(*
SPDX-FileCopyrightText: c 2026 Oleksandr Tiutyk <trofimich@gmail.com>
SPDX-License-Identifier: MIT
License: https://opensource.org/license/mit
*)

(*!
<summary>Checks trimming direction, custom characters and complete removal.</summary>
<description>
Uses one task and stays at a stable address while assertions are bound to this instance.
</description>
*)

{attribute 'no_assign'}
{attribute 'no_explicit_call' := 'do not call this function block directly'}
FUNCTION_BLOCK StringTrimTest EXTENDS TOF_Testing.SingleCycleTest
VAR_STAT
	{attribute 'hide'}
	_ClassName : STRING := __POUNAME();
END_VAR

(*!
<summary>Checks trimming direction, custom characters and complete removal.</summary>
*)
METHOD PROTECTED ExecuteTest
VAR
	text : STRING;
END_VAR
text := '  123   ';
TOF_Core.Strings.TrimChar(stringToTrim := text, trimMode := TOF_Core.TRIM_MODE.LEFT_AND_RIGHT);
Assert.ThatBool(
	actual := text = '123',
	message := "TrimChar must apply LEFT_AND_RIGHT exactly"
).IsTrue();

text := '  123   ';
TOF_Core.Strings.TrimChar(stringToTrim := text, trimMode := TOF_Core.TRIM_MODE.LEFT);
Assert.ThatBool(
	actual := text = '123   ',
	message := "TrimChar must apply LEFT exactly"
).IsTrue();

text := '  123   ';
TOF_Core.Strings.TrimChar(stringToTrim := text, trimMode := TOF_Core.TRIM_MODE.RIGHT);
Assert.ThatBool(
	actual := text = '  123',
	message := "TrimChar must apply RIGHT exactly"
).IsTrue();

text := '**a*b**';
TOF_Core.Strings.TrimChar(stringToTrim := text, trimMode := TOF_Core.TRIM_MODE.LEFT_AND_RIGHT, trimChar := '*');
Assert.ThatBool(
	actual := text = 'a*b',
	message := "Trimming a custom character must preserve an internal match"
).IsTrue();

text := '***';
TOF_Core.Strings.TrimChar(stringToTrim := text, trimChar := '*');
Assert.ThatBool(
	actual := text = '',
	message := "Trimming all matching characters must make the result empty"
).IsTrue();
END_METHOD

//! <summary>Borrows the concrete class name. Callers must not modify it.</summary>
{attribute 'monitoring' := 'call'}
PROPERTY ClassName : REFERENCE TO STRING
GET
ClassName REF= _ClassName;
END_GET
END_PROPERTY

//! <summary>Borrows the compiler-initialized namespace name. Callers must not modify it.</summary>
{attribute 'monitoring' := 'call'}
PROPERTY NamespaceName : REFERENCE TO STRING
GET
NamespaceName REF= CurrentNamespace.Name;
END_GET
END_PROPERTY

//! <summary>Reports the concrete instance size in bytes.</summary>
{attribute 'monitoring' := 'call'}
PROPERTY SelfSize : ULINT
GET
SelfSize := XSIZEOF(THIS^);
END_GET
END_PROPERTY

END_FUNCTION_BLOCK

(* stored: Version 1.1.0.1
   POU StringTrimTest: Id {87bf74ee-f5a5-4675-896e-b5ee7479797d}, SpecialFunc None
   Method ExecuteTest: Id {cb39fbf7-2963-4172-9d3a-4e67ed250509}
   Property ClassName: Id {ddcfa616-8518-4416-861a-835eac7ac173}
   Get Get: Id {5413b56c-7e0c-43e9-9d0b-e6d09ccb35cb}
   Property NamespaceName: Id {f6aafb92-d957-4bc6-a99e-56860fa12933}
   Get Get: Id {cfeb6518-bb70-4915-a35d-969e6f7ca66c}
   Property SelfSize: Id {ea725ccf-0d6a-4315-9ff6-fb4961a2156e}
   Get Get: Id {d3183065-bb3e-42e8-bdef-23f4b6e3f13d} *)
